// TIA Portal V21 export
// export: Created 2026-11-10T07:35:14.1141107Z, ExportSetting WithDefaults, DisplayName Totally Integrated Automation Portal, DisplayVersion V21 Update 3, DisplayName STEP 7 Professional, DisplayVersion V21 Update 3, DisplayName STEP 7 Safety, DisplayVersion V21, DisplayName Tech WebApplication, DisplayVersion V21, DisplayName WinCC Basic/Comfort/Advanced, DisplayVersion V21 Update 3, DisplayName WinCC Unified, DisplayVersion V21 Update 3
FUNCTION_BLOCK "FB_Lad_ex113"   // FB38, LAD
{ S7_Optimized_Access := 'TRUE' }
VERSION : 0.1
// stored: AutoNumber true, IsIECCheckEnabled false, IsRetainMemResEnabled false, MemoryReserve 100, SetENOAutomatically false, UDAEnableTagReadback false
   VAR_INPUT
      v_prgflt_reset_mask : DWord;
      v_accflt_reset_mask : DWord;
      v_ret_val : Int;
   END_VAR
   VAR_OUTPUT
      v_prgflt_masked : DWord;
      v_accflt_masked : DWord;
   END_VAR
BEGIN

REGION Network 1: DMSK_FLT - Unmask synchronous error events
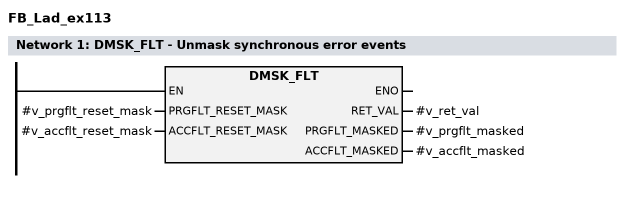
   RUNG wire#powerrail
      DMSK_FLT(PRGFLT_RESET_MASK := #v_prgflt_reset_mask, ACCFLT_RESET_MASK := #v_accflt_reset_mask, RET_VAL => #v_ret_val, PRGFLT_MASKED => #v_prgflt_masked, ACCFLT_MASKED => #v_accflt_masked)
   END_RUNG
   // the same network as SCL:
   #v_ret_val := DMSK_FLT(PRGFLT_RESET_MASK := #v_prgflt_reset_mask,
                          ACCFLT_RESET_MASK := #v_accflt_reset_mask,
                          PRGFLT_MASKED => #v_prgflt_masked,
                          ACCFLT_MASKED => #v_accflt_masked);
END_REGION
END_FUNCTION_BLOCK
